// TIA Portal V20 export
// export: Created 2026-10-11T05:28:41.0621708Z, ExportSetting WithDefaults, DisplayName Totally Integrated Automation Portal, DisplayVersion V20, DisplayName TIA Portal Openness, DisplayVersion V20, DisplayName TIA Portal Teamcenter Gateway, DisplayVersion V20, DisplayName TIA Portal Version Control Interface, DisplayVersion V20, DisplayName SINAMICS Startdrive Advanced, DisplayVersion V20 SP1 Update 2, DisplayName SINAMICS Startdrive G110M, G120, G120C, G120D, G120P, G115D, DisplayVersion V20 SP1 Update 2, DisplayName SINAMICS Startdrive G130, G150, S120, S150, SINAMICS MV, G220, S200, S210, DisplayVersion V20 SP1 Update 2, DisplayName STEP 7 Professional, DisplayVersion V20, DisplayName STEP 7 Safety, DisplayVersion V20, DisplayName WinCC Basic/Comfort/Advanced, DisplayVersion V20, DisplayName WinCC Professional, DisplayVersion V20, DisplayName WinCC Unified, DisplayVersion V20
FUNCTION "FRK_UnitFollow" : Void   // FC59, SCL
{ S7_Optimized_Access := 'TRUE' }
VERSION : 0.1
// stored: AutoNumber true, IsIECCheckEnabled false, SetENOAutomatically false, UDAEnableTagReadback false
   VAR_INPUT
      Supported : Array[0..6] of Bool;
   END_VAR
   VAR_IN_OUT
      Core : "FRK_Core";
      Unit : "FRK_Unit";
      Status : "ST_ModuleStatus";
      Policy : Array[0..6] of "ST_ModePolicy";
      Access : "FRK_Access";
   END_VAR
   VAR_TEMP
      Request : "ST_HmiRequest";
   END_VAR
BEGIN

   IF #Unit.FollowStart AND NOT #Unit.ModePending AND NOT #Unit.Clearing THEN
       #Unit.FollowStart := FALSE;
       #Request.Kind := 5;
       "FRK_UnitOperation"(Core := #Core,
                           Unit := #Unit,
                           Status := #Status,
                           Policy := #Policy,
                           Access := #Access,
                           Supported := #Supported,
                           Request := #Request,
                           Response := "FRK_UnitScratch".Response,
                           Trusted := TRUE);
   END_IF;
END_FUNCTION
